TYPE "ST_ReleaseReport"
VERSION : 0.1
   STRUCT
      Released : Bool;
      Count : Int;
      Reasons : Array[1..24] of "ST_ReleaseReason";
   END_STRUCT;

END_TYPE

